(* IEC 61131-3 sources: Codesys_IAP/Demo/PLC1/PLC 1 Simulatie Ladder StructuredTekst IOStructures 2V0_tekst/Programma Ladder, 6 files *)

(* ---- BedieningPrg.st ---- *)
(*#### DECLARATIE ####*)
PROGRAM BedieningPrg
VAR
END_VAR

(* ---- HoofdPrg.st ---- *)
(*#### DECLARATIE ####*)
PROGRAM HoofdPrg
VAR_INPUT
	// Reset het programma
	Px_HoofdReset: BOOL;
	// Start het programma
	Px_HoofdStart: BOOL;
	// Reset de SFC bv Noodstop
	SFCInit: BOOL;
END_VAR
VAR_OUTPUT
	// Er is een error op getreden
	Px_HoofdError: BOOL;
	// Commando is uitgevoerd
	Px_HoofdGereed: BOOL;
	// Programma is bezig
	Px_HoofdBezig: BOOL;
	// Programma is aan het opstarten
	Px_HoofdOpstart: BOOL;
END_VAR

(* ---- MagazijnPrg.st ---- *)
(*#### DECLARATIE ####*)
PROGRAM MagazijnPrg

VAR_INPUT
	// Reset het magazijn na start of error
	Px_MagazijnReset: BOOL;
	// Start uitstoten
	Px_MagazijnStart: BOOL;

	// Reset de SFC bv Noodstop
	SFCInit: BOOL;
	// Enable runtime limit checks
	SFCEnableLimit: BOOL := TRUE;
	// Reset runtime error
	SFCQuitError : BOOL;
END_VAR

VAR_OUTPUT
	// Er is een error opgetreden
	Px_MagazijnError: BOOL;
	// Commando is uitgevoerd
	Px_MagazijnGereed: BOOL;
	// Bezig met uitvoeren van commando
	Px_MagazijnBezig: BOOL;
	// Runtime limit is opgetreden
	SFCError: BOOL;
END_VAR

VAR
	// Tijdsvertraging voor fouten
	Mx_Error: BOOL;
END_VAR

(* ---- OverzetterPrg.st ---- *)
(*#### DECLARATIE ####*)
PROGRAM OverzetterPrg
VAR_INPUT
	// Reset de overzetter na start of error
	Px_OverzetterReset: BOOL;
	// Start de overzetter
	Px_OverzetterStart: BOOL;

	// Reset de SFC bv Noodstop
	SFCInit: BOOL;
	// Enable runtime limit checks
	SFCEnableLimit: BOOL := TRUE;
	// Reset runtime error
	SFCQuitError : BOOL;
END_VAR
VAR_OUTPUT
	// Overzetter heeft een error
	Px_OverzetterError: BOOL;
	// Overzetter heeft opdracht uitgevoerd
	Px_OverzetterGereed: BOOL;
	// Overzetter is bezig
	Px_OverzetterBezig: BOOL;
	// Runtime limit is opgetreden
	SFCError: BOOL;
END_VAR
VAR
	// Tijdsvertraging voor sommige stappen
	Mx_Delay: BOOL;
END_VAR

(* ---- SignaleringPrg.st ---- *)
(*#### DECLARATIE ####*)
PROGRAM SignaleringPrg
VAR
	// Knipperen gele lamp
	Fb_GeelKnipper: Blink;
END_VAR

(* ---- SorterenPrg.st ---- *)
(*#### DECLARATIE ####*)
PROGRAM SorterenPrg
VAR_INPUT
	// Reset de sorteren na start of error
	Px_SorterenReset: BOOL;
	// Start het sorteren
	Px_SorterenStart: BOOL;

	// Reset de SFC bv Noodstop
	SFCInit: BOOL;
	// Enable runtime limit checks
	SFCEnableLimit: BOOL := TRUE;
	// Reset runtime error
	SFCQuitError : BOOL;
END_VAR
VAR_OUTPUT
	// Sorteren heeft een error
	Px_SorterenError: BOOL;
	// Sorteren heeft een opdracht uitgevoerd
	Px_SorterenGereed: BOOL;
	// Sorteren is bezig
	Px_SorterenBezig: BOOL;
	// Runtime limit is opgetreden
	SFCError: BOOL;
END_VAR
